(* Schneider Machine Expert - Basic project Projeto Charpy 3 - Prático V1, file version 3.0.0.0 *)
(* ProjectInformations: Name=Novo projeto *)

HARDWARE
  Cpu 0: TM221CE40R
  EthernetConfiguration: NetworkName=M221, IpAllocationMode=FixedAddress, IpAddress=10.0.0.20, SubnetMask=255.0.0.0
  SerialLineConfiguration: Baud=Baud19200, Parity=ParityEven, DataBits=DataBits8, StopBits=StopBits1, PhysicalMedium=PhysicalMediumRs485, TransmissionMode=TransmissionModeModbusRtu, SlaveId=1, Addressing=SlaveAddressing
  MastTask: UsePeriodScanMode=false, PeriodScan=100
  FastTask: Period=255
  CpuBehavior: StartingMode=StartAsPreviousState, AutoSaveRamOnEeprom=true, WatchdogPeriod=250

SYMBOLS  (address, symbol, comment, settings)
  %HSC0.V   VALOR_ENCODER  "Entrada de alta velocidade"
  %M0         "Engrenagem"
  %M1         "Motor Subir"
  %M2         "Motor Descer"
  %M3         "Impacto"
  %M5         "Perdas"
  %M6         "Perdas_aux"
  %M7         "Aux_subir"
  %M20        "ATRITO_OK"
  %M21        "ATRITO_FALHO"
  %M31      SENSOR_VIRTUAL_B  "Virtual_Baixo"
  %M32      SENSOR_VIRTUAL_C  "Virtual_Cima"
  %S6       SB_TB1S  "Base de tempo de 1 s gerada por um relógio interno"
  %MW0      PULSOS_ENCODER  "Pulsos brutos do encoder"
  %MF2      ANGULO_ATUAL  "Ângulo instantâneo em Graus"
  %MF4      ANGULO_PICO  "Maior ângulo atingido no impacto"
  %MF6      ENERGIA_NOMINAL  "Capacidade da ponta do martelo"
  %MF8      ENERGIA_ABSORVIDA  "Resultado final do ensaio em Joules"
  %MF10     MF_10
  %MF12     MF_12
  %MF120    PERDAS_J  "Energia perdida por atrito em Joules"
  %TM0        [Type=TP, Preset=75, Base=OneHundredMilliSeconds]
  %TM1        [Type=TP, Preset=75, Base=OneHundredMilliSeconds]
  %TM2        [Type=TP, Preset=1, Base=OneSecond]
  %TM3        [Type=TP, Preset=1, Base=OneSecond]
  %TM4        [Type=TP, Preset=60, Base=OneSecond]
  %TM6        [Preset=15, Base=TenMilliSeconds]
  %TM7        [Preset=15, Base=TenMilliSeconds]
  %TM8        [Preset=15, Base=TenMilliSeconds]
  %I0.2     BOT_RESET  "Botão físico de zerar encoder e pico"
  %I0.10    SENSOR_PORTA  "Sensor se a porta está fechada"
  %I0.11    SENSOR_BAIXO  "Sensor se o braço está em baixo"
  %I0.12    SENSOR_CIMA  "Sensor se o braço está em cima"
  %I0.19    BOTÃO_ATRITO  "Botão que inicia o teste de atrito"
  %I0.20    BOTÃO_ZERAR  "Botão que zera a referência do encoder"
  %I0.21    BOTÃO_IMPACTO  "Botão que libera para o impacto"
  %I0.22    BOTÃO_DESCER  "Botão que aciona por 7s"
  %I0.23    BOTÃO_SUBIR  "Botão que aciona por 7s"
  %Q0.0     Q_0_0  "Encaixe Engrenagem"
  %Q0.1     Q_0_1  "Motor Subir"
  %Q0.2     Q_0_2  "Motor Descer"
  %Q0.3     Q_0_3  "Liberar Catraca"
  %Q0.4     Q_0_4  "Liga Esteira"
  %Q0.5     Q_0_5  "Led Porta"
  %Q0.14    Q_0_14
  %Q0.15    Q_0_15
  %IW0.0    IN_ANALOG  "Valor do Potenciômetro"  [Type=Type_0_10V, Scope=Scope_Normal, Minimum=0, Maximum=1000]
  %HSC0       [Type=CounterOrDownCounterBiPhasesX4, Preset=0, DedicatedInputs(DedicatedInput(Activated=true), DedicatedInput(Activated=true)), ReflexOutputs(ReflexOutput(Activated=false, LessThanS0=false, GreaterOrEqualThanS0=false, GreaterOrEqualThanS1=false), ReflexOutput(Activated=false, LessThanS0=false, GreaterOrEqualThanS0=false, GreaterOrEqualThanS1=false)), Thresholds(Threshold(ThresholdType=NotUsed, Pri]

POU Novo POU
  (* SectionNumber=1 *)

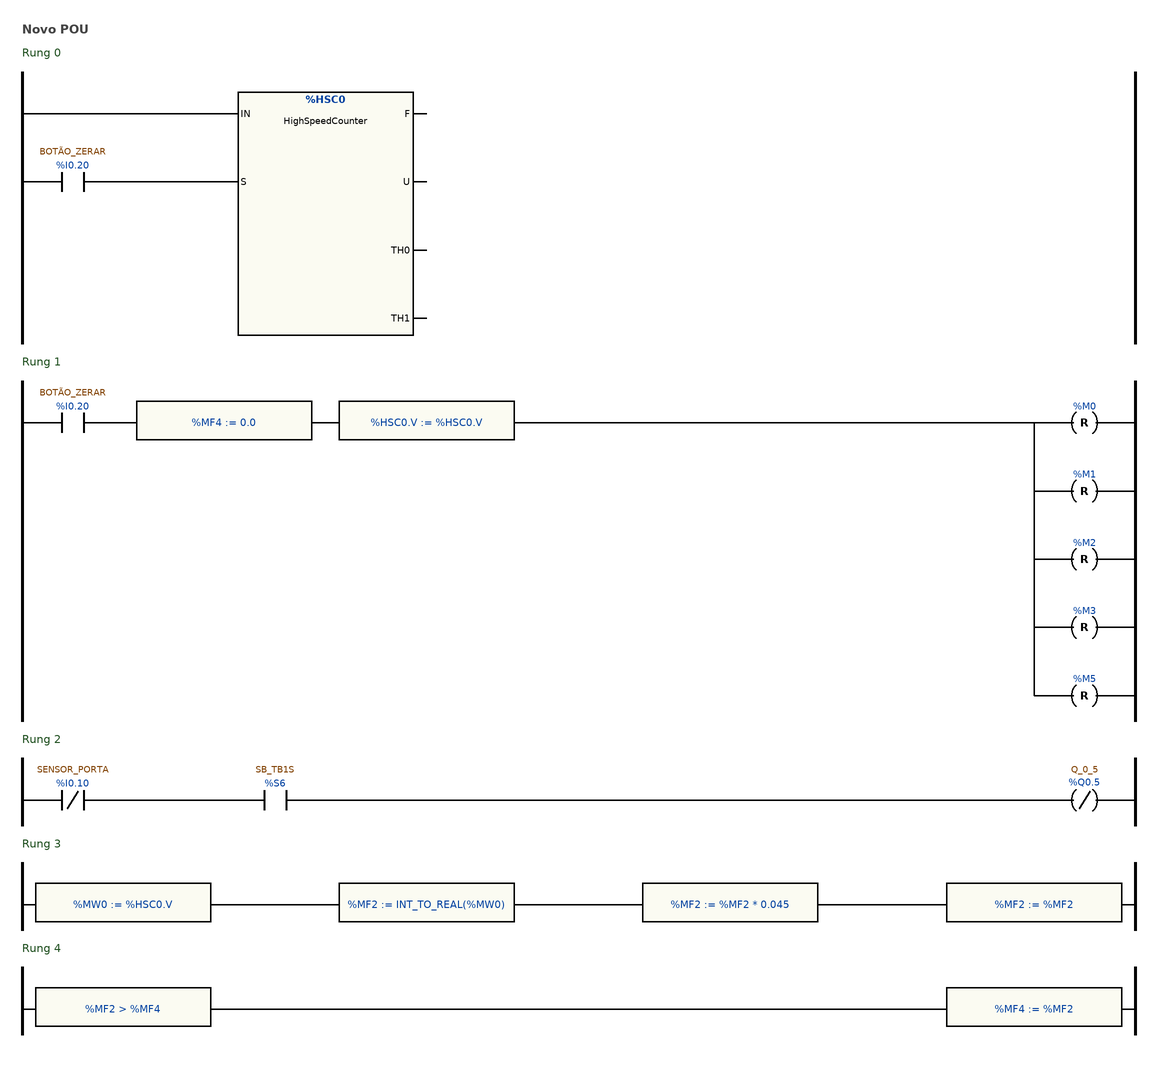

// Rung 0
  BLK %HSC0
  LD 1
  IN
  LD %I0.20               (* BOTÃO_ZERAR *)
  S
  END_BLK
  // as ST:
  //   %HSC0(IN := TRUE, S := BOTÃO_ZERAR);

// Rung 1
  LD %I0.20               (* BOTÃO_ZERAR *)
  OPER [ %MF4 := 0.0 ]    (* ANGULO_PICO *)
  OPER [ %HSC0.V := %HSC0.V ]
  R %M0
  R %M1
  R %M2
  R %M3
  R %M5
  // as ST:
  //   IF BOTÃO_ZERAR THEN ANGULO_PICO := 0.0; END_IF;
  //   IF BOTÃO_ZERAR THEN %HSC0.V := %HSC0.V; END_IF;
  //   IF BOTÃO_ZERAR THEN %M0 := FALSE; END_IF;
  //   IF BOTÃO_ZERAR THEN %M1 := FALSE; END_IF;
  //   IF BOTÃO_ZERAR THEN %M2 := FALSE; END_IF;
  //   IF BOTÃO_ZERAR THEN %M3 := FALSE; END_IF;
  //   IF BOTÃO_ZERAR THEN %M5 := FALSE; END_IF;

// Rung 2
  LDN %I0.10              (* SENSOR_PORTA *)
  AND %S6                 (* SB_TB1S *)
  STN %Q0.5               (* Q_0_5 *)
  // as ST:
  //   Q_0_5 := NOT (NOT SENSOR_PORTA AND SB_TB1S);

// Rung 3
  LD 1
  OPER [ %MW0 := %HSC0.V ](* PULSOS_ENCODER *)
  OPER [ %MF2 := INT_TO_REAL ( %MW0 ) ](* ANGULO_ATUAL, PULSOS_ENCODER *)
  OPER [ %MF2 := %MF2 * 0.045 ](* ANGULO_ATUAL, ANGULO_ATUAL *)
  [ %MF2 := %MF2 ]        (* ANGULO_ATUAL, ANGULO_ATUAL *)
  // as ST:
  //   PULSOS_ENCODER := %HSC0.V;
  //   ANGULO_ATUAL := INT_TO_REAL ( PULSOS_ENCODER );
  //   ANGULO_ATUAL := ANGULO_ATUAL * 0.045;
  //   ANGULO_ATUAL := ANGULO_ATUAL;

// Rung 4
  LD [ %MF2 > %MF4 ]      (* ANGULO_ATUAL, ANGULO_PICO *)
  [ %MF4 := %MF2 ]        (* ANGULO_PICO, ANGULO_ATUAL *)
  // as ST:
  //   IF ANGULO_ATUAL > ANGULO_PICO THEN ANGULO_PICO := ANGULO_ATUAL; END_IF;

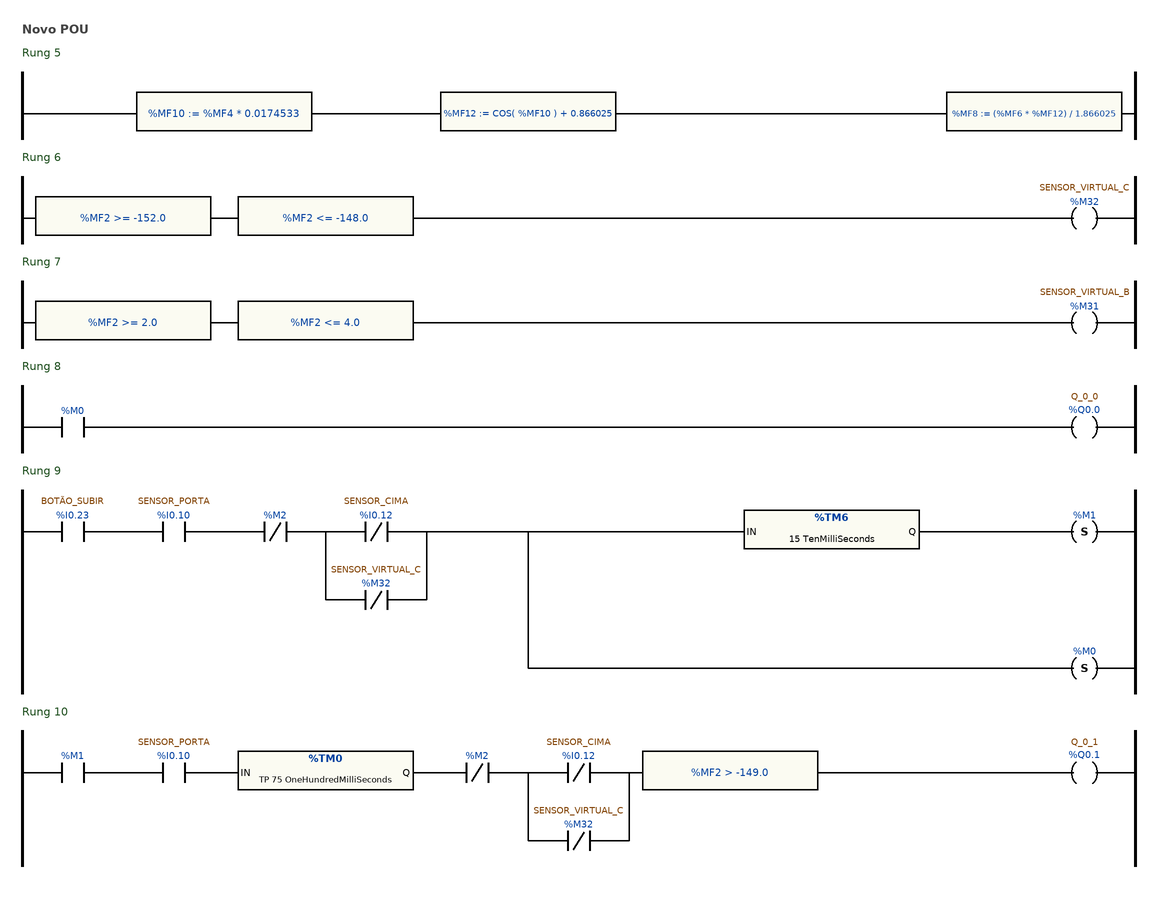

// Rung 5
  LD 1
  OPER [ %MF10 := %MF4 * 0.0174533 ](* MF_10, ANGULO_PICO *)
  OPER [ %MF12 := COS ( %MF10 ) + 0.866025 ](* MF_12, MF_10 *)
  [ %MF8 := ( %MF6 * %MF12 ) / 1.866025 ](* ENERGIA_ABSORVIDA, ENERGIA_NOMINAL, MF_12 *)
  // as ST:
  //   MF_10 := ANGULO_PICO * 0.0174533;
  //   MF_12 := COS ( MF_10 ) + 0.866025;
  //   ENERGIA_ABSORVIDA := ( ENERGIA_NOMINAL * MF_12 ) / 1.866025;

// Rung 6
  LD [ %MF2 >= -152.0 ]   (* ANGULO_ATUAL *)
  AND [ %MF2 <= -148.0 ]  (* ANGULO_ATUAL *)
  ST %M32                 (* SENSOR_VIRTUAL_C *)
  // as ST:
  //   SENSOR_VIRTUAL_C := ANGULO_ATUAL >= -152.0 AND ANGULO_ATUAL <= -148.0;

// Rung 7
  LD [ %MF2 >= 2.0 ]      (* ANGULO_ATUAL *)
  AND [ %MF2 <= 4.0 ]     (* ANGULO_ATUAL *)
  ST %M31                 (* SENSOR_VIRTUAL_B *)
  // as ST:
  //   SENSOR_VIRTUAL_B := ANGULO_ATUAL >= 2.0 AND ANGULO_ATUAL <= 4.0;

// Rung 8
  LD %M0
  ST %Q0.0                (* Q_0_0 *)
  // as ST:
  //   Q_0_0 := %M0;

// Rung 9
  LD 1
  MULTIFB
  LD 1
  AND %I0.23              (* BOTÃO_SUBIR *)
  AND %I0.10              (* SENSOR_PORTA *)
  ANDN %M2
  AND(N %I0.12            (* SENSOR_CIMA *)
  ORN %M32                (* SENSOR_VIRTUAL_C *)
  )
  ST %MW2009:X0
  BLK %TM6
  LD %MW2009:X0
  IN
  OUT_BLK
  LD Q
  S %M1
  END_BLK
  LD %MW2009:X0
  S %M0
  MULTIFB
  // as ST:
  //   %TM6(IN := BOTÃO_SUBIR AND SENSOR_PORTA AND NOT %M2 AND (NOT SENSOR_CIMA OR NOT SENSOR_VIRTUAL_C));
  //   IF %TM6.Q THEN %M1 := TRUE; END_IF;
  //   IF BOTÃO_SUBIR AND SENSOR_PORTA AND NOT %M2 AND (NOT SENSOR_CIMA OR NOT SENSOR_VIRTUAL_C) THEN %M0 := TRUE; END_IF;

// Rung 10
  BLK %TM0
  LD %M1
  AND %I0.10              (* SENSOR_PORTA *)
  IN
  OUT_BLK
  LD Q
  ANDN %M2
  AND(N %I0.12            (* SENSOR_CIMA *)
  ORN %M32                (* SENSOR_VIRTUAL_C *)
  )
  AND [ %MF2 > -149.0 ]   (* ANGULO_ATUAL *)
  ST %Q0.1                (* Q_0_1 *)
  END_BLK
  // as ST:
  //   %TM0(IN := %M1 AND SENSOR_PORTA);
  //   Q_0_1 := %TM0.Q AND NOT %M2 AND (NOT SENSOR_CIMA OR NOT SENSOR_VIRTUAL_C) AND ANGULO_ATUAL > -149.0;

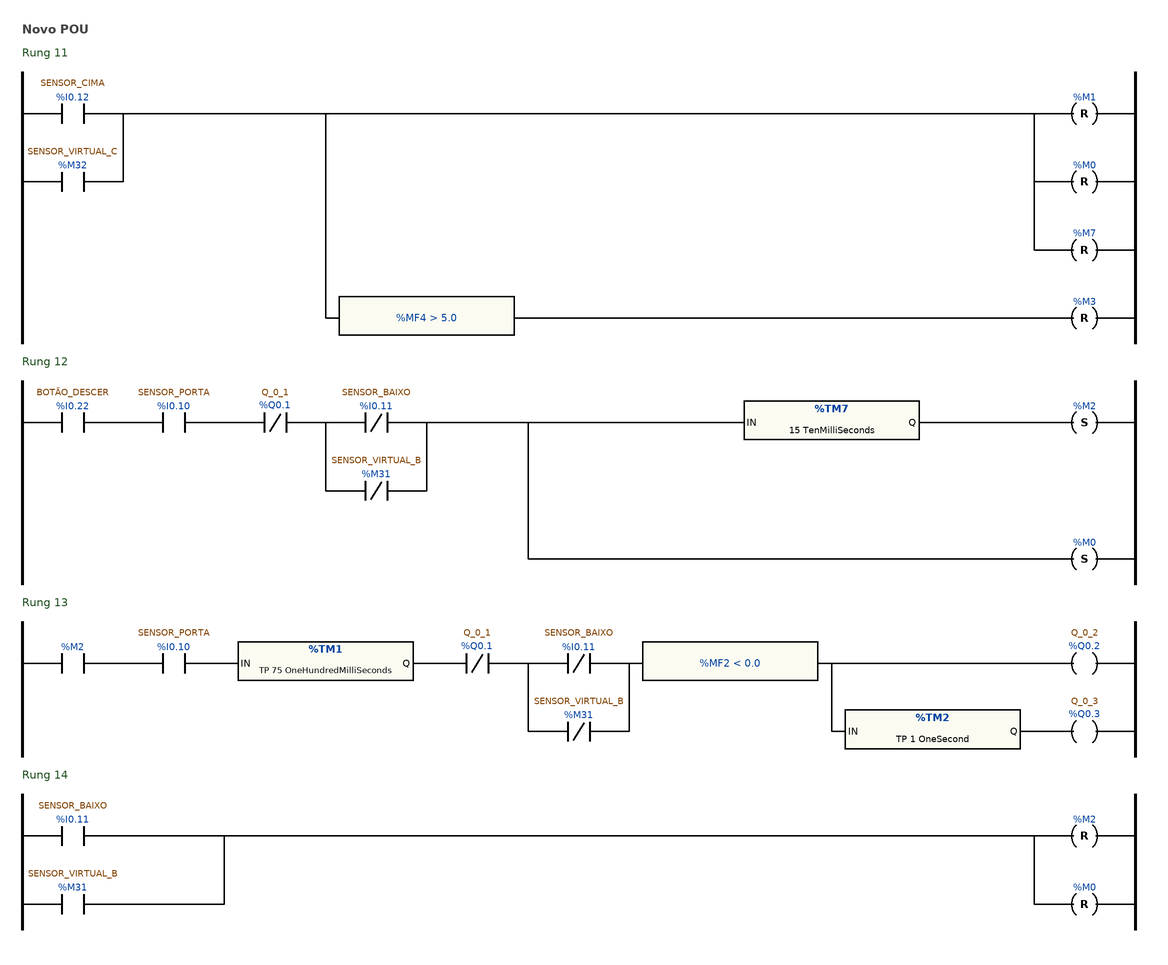

// Rung 11
  LD %I0.12               (* SENSOR_CIMA *)
  OR %M32                 (* SENSOR_VIRTUAL_C *)
  MPS
  R %M1
  R %M0
  R %M7
  MPP
  AND [ %MF4 > 5.0 ]      (* ANGULO_PICO *)
  R %M3
  // as ST:
  //   IF SENSOR_CIMA OR SENSOR_VIRTUAL_C THEN %M1 := FALSE; END_IF;
  //   IF SENSOR_CIMA OR SENSOR_VIRTUAL_C THEN %M0 := FALSE; END_IF;
  //   IF SENSOR_CIMA OR SENSOR_VIRTUAL_C THEN %M7 := FALSE; END_IF;
  //   IF (SENSOR_CIMA OR SENSOR_VIRTUAL_C) AND ANGULO_PICO > 5.0 THEN %M3 := FALSE; END_IF;

// Rung 12
  LD 1
  MULTIFB
  LD 1
  AND %I0.22              (* BOTÃO_DESCER *)
  AND %I0.10              (* SENSOR_PORTA *)
  ANDN %Q0.1              (* Q_0_1 *)
  AND(N %I0.11            (* SENSOR_BAIXO *)
  ORN %M31                (* SENSOR_VIRTUAL_B *)
  )
  ST %MW2009:X0
  BLK %TM7
  LD %MW2009:X0
  IN
  OUT_BLK
  LD Q
  S %M2
  END_BLK
  LD %MW2009:X0
  S %M0
  MULTIFB
  // as ST:
  //   %TM7(IN := BOTÃO_DESCER AND SENSOR_PORTA AND NOT Q_0_1 AND (NOT SENSOR_BAIXO OR NOT SENSOR_VIRTUAL_B));
  //   IF %TM7.Q THEN %M2 := TRUE; END_IF;
  //   IF BOTÃO_DESCER AND SENSOR_PORTA AND NOT Q_0_1 AND (NOT SENSOR_BAIXO OR NOT SENSOR_VIRTUAL_B) THEN %M0 := TRUE; END_IF;

// Rung 13
  LD 1
  MULTIFB
  BLK %TM1
  LD 1
  AND %M2
  AND %I0.10              (* SENSOR_PORTA *)
  IN
  OUT_BLK
  LD Q
  ST %MW2009:X0
  END_BLK
  LD %MW2009:X0
  ANDN %Q0.1              (* Q_0_1 *)
  AND(N %I0.11            (* SENSOR_BAIXO *)
  ORN %M31                (* SENSOR_VIRTUAL_B *)
  )
  AND [ %MF2 < 0.0 ]      (* ANGULO_ATUAL *)
  ST %MW2009:X1
  LD %MW2009:X1
  ST %Q0.2                (* Q_0_2 *)
  BLK %TM2
  LD %MW2009:X1
  IN
  OUT_BLK
  LD Q
  ST %Q0.3                (* Q_0_3 *)
  END_BLK
  MULTIFB
  // as ST:
  //   %TM1(IN := %M2 AND SENSOR_PORTA);
  //   Q_0_2 := %TM1.Q AND NOT Q_0_1 AND (NOT SENSOR_BAIXO OR NOT SENSOR_VIRTUAL_B) AND ANGULO_ATUAL < 0.0;
  //   %TM2(IN := %TM1.Q AND NOT Q_0_1 AND (NOT SENSOR_BAIXO OR NOT SENSOR_VIRTUAL_B) AND ANGULO_ATUAL < 0.0);
  //   Q_0_3 := %TM2.Q;

// Rung 14
  LD %I0.11               (* SENSOR_BAIXO *)
  OR %M31                 (* SENSOR_VIRTUAL_B *)
  R %M2
  R %M0
  // as ST:
  //   IF SENSOR_BAIXO OR SENSOR_VIRTUAL_B THEN %M2 := FALSE; END_IF;
  //   IF SENSOR_BAIXO OR SENSOR_VIRTUAL_B THEN %M0 := FALSE; END_IF;

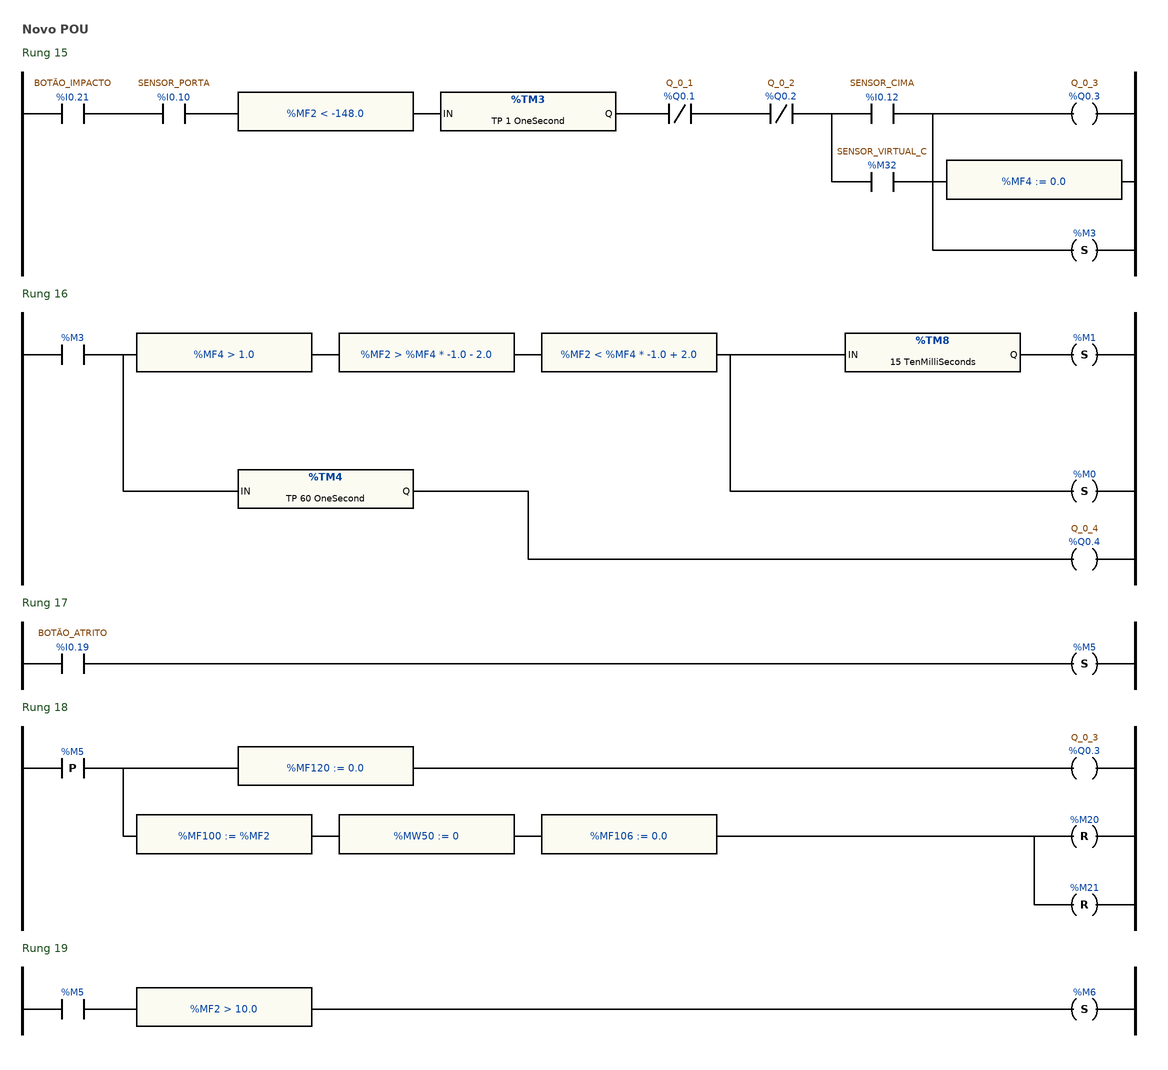

// Rung 15
  BLK %TM3
  LD %I0.21               (* BOTÃO_IMPACTO *)
  AND %I0.10              (* SENSOR_PORTA *)
  AND [ %MF2 < -148.0 ]   (* ANGULO_ATUAL *)
  IN
  OUT_BLK
  LD Q
  ANDN %Q0.1              (* Q_0_1 *)
  ANDN %Q0.2              (* Q_0_2 *)
  AND( %I0.12             (* SENSOR_CIMA *)
  OR %M32                 (* SENSOR_VIRTUAL_C *)
  )
  ST %Q0.3                (* Q_0_3 *)
  [ %MF4 := 0.0 ]         (* ANGULO_PICO *)
  S %M3
  END_BLK
  // as ST:
  //   %TM3(IN := BOTÃO_IMPACTO AND SENSOR_PORTA AND ANGULO_ATUAL < -148.0);
  //   Q_0_3 := %TM3.Q AND NOT Q_0_1 AND NOT Q_0_2 AND (SENSOR_CIMA OR SENSOR_VIRTUAL_C);
  //   IF %TM3.Q AND NOT Q_0_1 AND NOT Q_0_2 AND (SENSOR_CIMA OR SENSOR_VIRTUAL_C) THEN ANGULO_PICO := 0.0; END_IF;
  //   IF %TM3.Q AND NOT Q_0_1 AND NOT Q_0_2 AND (SENSOR_CIMA OR SENSOR_VIRTUAL_C) THEN %M3 := TRUE; END_IF;

// Rung 16
  LD 1
  MULTIFB
  LD 1
  AND %M3
  ST %MW2009:X0
  LD %MW2009:X0
  AND [ %MF4 > 1.0 ]      (* ANGULO_PICO *)
  AND [ %MF2 > %MF4 * -1.0 - 2.0 ](* ANGULO_ATUAL, ANGULO_PICO *)
  AND [ %MF2 < %MF4 * -1.0 + 2.0 ](* ANGULO_ATUAL, ANGULO_PICO *)
  ST %MW2009:X1
  BLK %TM8
  LD %MW2009:X1
  IN
  OUT_BLK
  LD Q
  S %M1
  END_BLK
  LD %MW2009:X1
  S %M0
  BLK %TM4
  LD %MW2009:X0
  IN
  OUT_BLK
  LD Q
  ST %Q0.4                (* Q_0_4 *)
  END_BLK
  MULTIFB
  // as ST:
  //   %TM8(IN := %M3 AND ANGULO_PICO > 1.0 AND ANGULO_ATUAL > ANGULO_PICO * -1.0 - 2.0 AND ANGULO_ATUAL < ANGULO_PICO * -1.0 + 2.0);
  //   IF %TM8.Q THEN %M1 := TRUE; END_IF;
  //   IF %M3 AND ANGULO_PICO > 1.0 AND ANGULO_ATUAL > ANGULO_PICO * -1.0 - 2.0 AND ANGULO_ATUAL < ANGULO_PICO * -1.0 + 2.0 THEN %M0 := TRUE; END_IF;
  //   %TM4(IN := %M3);
  //   Q_0_4 := %TM4.Q;

// Rung 17
  LD %I0.19               (* BOTÃO_ATRITO *)
  S %M5
  // as ST:
  //   IF BOTÃO_ATRITO THEN %M5 := TRUE; END_IF;

// Rung 18
  LDR %M5
  MPS
  OPER [ %MF120 := 0.0 ]  (* PERDAS_J *)
  ST %Q0.3                (* Q_0_3 *)
  MPP
  OPER [ %MF100 := %MF2 ] (* ANGULO_ATUAL *)
  OPER [ %MW50 := 0 ]
  OPER [ %MF106 := 0.0 ]
  R %M20
  R %M21
  // as ST:
  //   IF RISING(%M5) THEN PERDAS_J := 0.0; END_IF;
  //   Q_0_3 := RISING(%M5);
  //   IF RISING(%M5) THEN %MF100 := ANGULO_ATUAL; END_IF;
  //   IF RISING(%M5) THEN %MW50 := 0; END_IF;
  //   IF RISING(%M5) THEN %MF106 := 0.0; END_IF;
  //   IF RISING(%M5) THEN %M20 := FALSE; END_IF;
  //   IF RISING(%M5) THEN %M21 := FALSE; END_IF;

// Rung 19
  LD %M5
  AND [ %MF2 > 10.0 ]     (* ANGULO_ATUAL *)
  S %M6
  // as ST:
  //   IF %M5 AND ANGULO_ATUAL > 10.0 THEN %M6 := TRUE; END_IF;

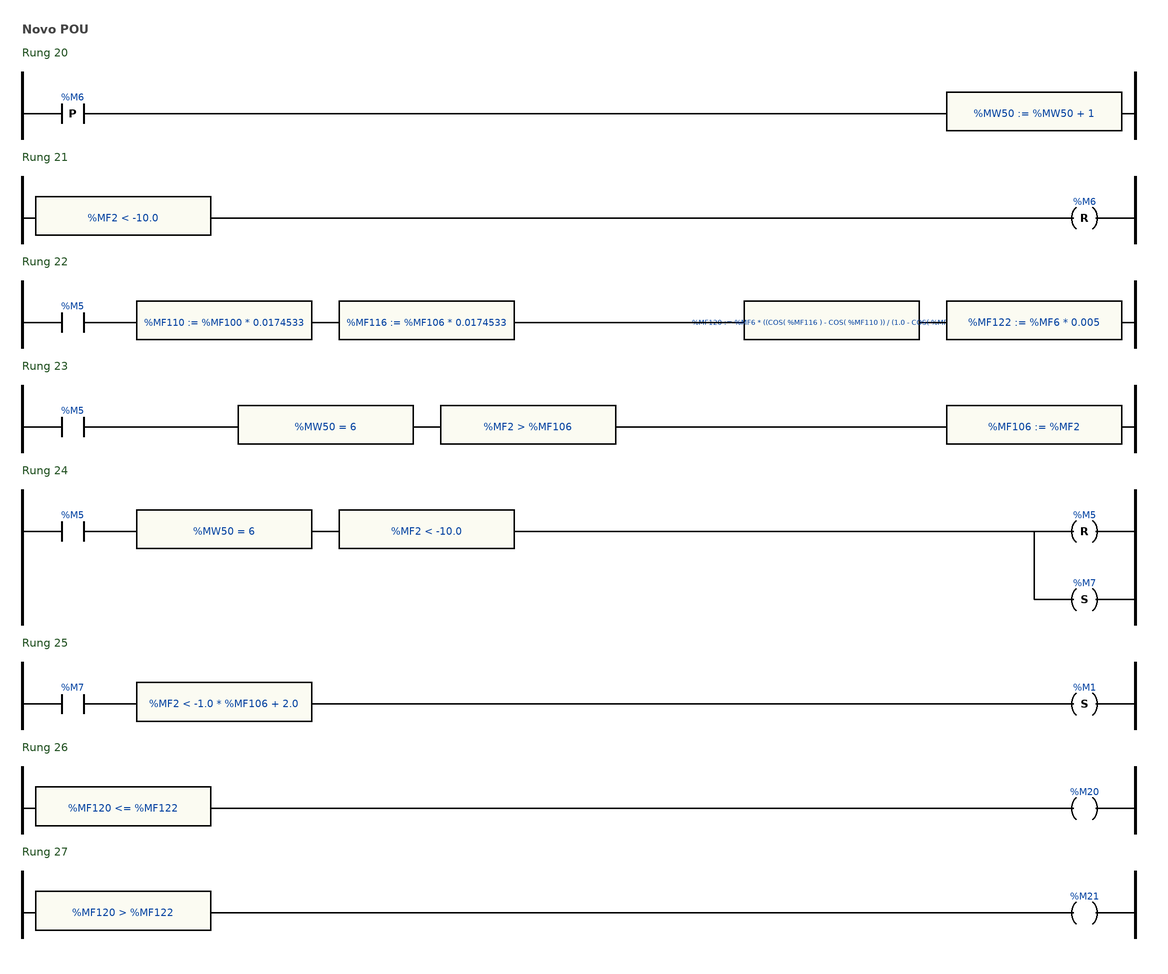

// Rung 20
  LDR %M6
  [ %MW50 := %MW50 + 1 ]
  // as ST:
  //   IF RISING(%M6) THEN %MW50 := %MW50 + 1; END_IF;

// Rung 21
  LD [ %MF2 < -10.0 ]     (* ANGULO_ATUAL *)
  R %M6
  // as ST:
  //   IF ANGULO_ATUAL < -10.0 THEN %M6 := FALSE; END_IF;

// Rung 22
  LD %M5
  OPER [ %MF110 := %MF100 * 0.0174533 ]
  OPER [ %MF116 := %MF106 * 0.0174533 ]
  OPER [ %MF120 := %MF6 * ( ( COS ( %MF116 ) - COS ( %MF110 ) ) / ( 1.0 - COS ( %MF110 ) ) ) ](* PERDAS_J, ENERGIA_NOMINAL *)
  [ %MF122 := %MF6 * 0.005 ](* ENERGIA_NOMINAL *)
  // as ST:
  //   IF %M5 THEN %MF110 := %MF100 * 0.0174533; END_IF;
  //   IF %M5 THEN %MF116 := %MF106 * 0.0174533; END_IF;
  //   IF %M5 THEN PERDAS_J := ENERGIA_NOMINAL * ( ( COS ( %MF116 ) - COS ( %MF110 ) ) / ( 1.0 - COS ( %MF110 ) ) ); END_IF;
  //   IF %M5 THEN %MF122 := ENERGIA_NOMINAL * 0.005; END_IF;

// Rung 23
  LD %M5
  AND [ %MW50 = 6 ]
  AND [ %MF2 > %MF106 ]   (* ANGULO_ATUAL *)
  [ %MF106 := %MF2 ]      (* ANGULO_ATUAL *)
  // as ST:
  //   IF %M5 AND %MW50 = 6 AND ANGULO_ATUAL > %MF106 THEN %MF106 := ANGULO_ATUAL; END_IF;

// Rung 24
  LD %M5
  AND [ %MW50 = 6 ]
  AND [ %MF2 < -10.0 ]    (* ANGULO_ATUAL *)
  R %M5
  S %M7
  // as ST:
  //   _t1 := %M5 AND %MW50 = 6 AND ANGULO_ATUAL < -10.0;
  //   IF _t1 THEN %M5 := FALSE; END_IF;
  //   IF _t1 THEN %M7 := TRUE; END_IF;

// Rung 25
  LD %M7
  AND [ %MF2 < -1.0 * %MF106 + 2.0 ](* ANGULO_ATUAL *)
  S %M1
  // as ST:
  //   IF %M7 AND ANGULO_ATUAL < -1.0 * %MF106 + 2.0 THEN %M1 := TRUE; END_IF;

// Rung 26
  LD [ %MF120 <= %MF122 ] (* PERDAS_J *)
  ST %M20
  // as ST:
  //   %M20 := PERDAS_J <= %MF122;

// Rung 27
  LD [ %MF120 > %MF122 ]  (* PERDAS_J *)
  ST %M21
  // as ST:
  //   %M21 := PERDAS_J > %MF122;
